(*
SPDX-FileCopyrightText: c 2026 Oleksandr Tiutyk <trofimich@gmail.com>
SPDX-License-Identifier: MIT
License: https://opensource.org/license/mit
*)

(*!
<summary>Checks strict and Try appends, including empty fragments and capacity failure.</summary>
<description>
Uses one task and stays at a stable address while assertions are bound to this instance.
</description>
*)

{attribute 'no_assign'}
{attribute 'no_explicit_call' := 'do not call this function block directly'}
FUNCTION_BLOCK StringAppendTest EXTENDS TOF_Testing.SingleCycleTest
VAR_STAT
	{attribute 'hide'}
	_ClassName : STRING := __POUNAME();
END_VAR

(*!
<summary>Checks strict and Try appends, including empty fragments and capacity failure.</summary>
<description>
Uses an eight-byte ASCII target. After a later fragment fails to fit, checks that the original text and the
first appended fragment remain at the start of the target.
</description>
*)
METHOD PROTECTED ExecuteTest
VAR
	target : STRING(8);
	accepted : BOOL;
	prefixFound : BOOL;
	prefixPosition : UDINT;
END_VAR
target := 'ab';
TOF_Core.Strings.Append255(target, 'cd', '', 'efgh');
Assert.ThatBool(
	actual := target = 'abcdefgh',
	message := "Append255 must skip an empty fragment and fill the target exactly"
).IsTrue();

target := 'ab';
accepted := TOF_Core.Strings.TryAppend255(
	targetString := target,
	sourceString1 := 'cd',
	sourceString2 := '',
	sourceString3 := 'efgh'
);
Assert.ThatBool(
	actual := accepted AND_THEN target = 'abcdefgh',
	message := "TryAppend255 must accept an exact fit"
).IsTrue();

target := 'ab';
accepted := TOF_Core.Strings.TryAppend255(
	targetString := target,
	sourceString1 := 'cd',
	sourceString2 := 'ABCDE',
	sourceString3 := '!'
);
Assert.ThatBool(
	actual := accepted,
	message := "TryAppend255 must report capacity failure"
).IsFalse();

prefixFound := TOF_Core.Strings.Find(
	stringToSearchIn := target,
	stringToFind := 'abcd',
	position => prefixPosition
);
Assert.ThatBool(
	actual := prefixFound AND_THEN prefixPosition = 1,
	message := "TryAppend255 must preserve the successfully appended prefix"
).IsTrue();

target := 'ab';
TOF_Core.Strings.Append(targetString := target, sourceString := 'cd');
TOF_Core.Strings.Append(targetString := target, sourceString := '');
TOF_Core.Strings.Append(targetString := target, sourceString := 'efgh');
Assert.ThatBool(
	actual := target = 'abcdefgh',
	message := "Append must preserve the target on empty input and accept the exact fit"
).IsTrue();

target := 'abcdef';
accepted := TOF_Core.Strings.TryAppend(targetString := target, sourceString := 'gh');
Assert.ThatBool(
	actual := accepted AND_THEN target = 'abcdefgh',
	message := "TryAppend must accept an exact fit"
).IsTrue();

accepted := TOF_Core.Strings.TryAppend(targetString := target, sourceString := 'i');
Assert.ThatBool(
	actual := accepted,
	message := "TryAppend must reject another character in a full target"
).IsFalse();
Assert.ThatBool(
	actual := target = 'abcdefgh',
	message := "TryAppend must preserve the full target when one more character does not fit"
).IsTrue();
END_METHOD

//! <summary>Borrows the concrete class name. Callers must not modify it.</summary>
{attribute 'monitoring' := 'call'}
PROPERTY ClassName : REFERENCE TO STRING
GET
ClassName REF= _ClassName;
END_GET
END_PROPERTY

//! <summary>Borrows the compiler-initialized namespace name. Callers must not modify it.</summary>
{attribute 'monitoring' := 'call'}
PROPERTY NamespaceName : REFERENCE TO STRING
GET
NamespaceName REF= CurrentNamespace.Name;
END_GET
END_PROPERTY

//! <summary>Reports the concrete instance size in bytes.</summary>
{attribute 'monitoring' := 'call'}
PROPERTY SelfSize : ULINT
GET
SelfSize := XSIZEOF(THIS^);
END_GET
END_PROPERTY

END_FUNCTION_BLOCK

(* stored: Version 1.1.0.1
   POU StringAppendTest: Id {db03c086-1446-4de2-8420-bf576b238b8c}, SpecialFunc None
   Method ExecuteTest: Id {52a3ca7e-de6e-4771-a459-227b72a987e4}
   Property ClassName: Id {43018df9-5ace-4511-9939-fe3f63f12018}
   Get Get: Id {782e7624-d488-4e97-967f-056f381b36dc}
   Property NamespaceName: Id {57f7ef22-c1cb-4e59-8ef0-73a9b32fe5f0}
   Get Get: Id {78920eb4-5554-4e37-a395-f228ecf5e622}
   Property SelfSize: Id {fdee6cd9-0eab-4b38-9ff6-a7defd216334}
   Get Get: Id {0a6dc22a-1bab-44b1-9bee-18f99a192902} *)
